Fanuc KAREL source: kt00718.KL

-- PROVISIONAL review KL for V940-1; original PC SHA256 199eca4cacc04294e224a3000934cf67fd7c4e2a3afa222573561e05f22a253b
-- Incomplete behavior may be omitted. Consult companion uncertainty JSON. Do not deploy.
PROGRAM KT00718
%NOLOCKGROUP
VAR
  OUT : BOOLEAN
-- UNRESOLVED_DECL P1 type=000101
-- UNRESOLVED_DECL P2 type=000101
BEGIN
  -- V9_ZERO_TABLE_METADATA_HINT layout=0001; no indexed target words; source/name/runtime held
  -- UNRESOLVED_PC offsets 5-20; opcodes 22,63,23
  -- UNRESOLVED_PC offsets 25-29; opcodes 7F
END KT00718
